// Mock of the hydraulics unit, which is both the brake (I_Brake) and the hydraulics (I_Hydraulics) on MONETS/MONETN.
// The Az/El brake is hydraulic and locks by itself without pressure: Enable := FALSE (hydraulics off) closes the brake, and after
// InjectPressureLoss() the brake is locked and OpenBrake() has no effect until Reset(). Nobody sets Enable TRUE in the rig, so the
// brake opens as before as long as the pressure is there (OpenBrake does not need Enable).
// A close wins over the opening in the same scan, as in HalfBROT FB_HydraulicsControl (a pending bCloseBrake clears bOpenBrake): after
// CloseBrake() an OpenBrake() has no effect until the body has run (the rig calls it at the end of the scan). MONETcommon#272: the
// enabled elevation requests the opening in every scan, after the telescope.
FUNCTION_BLOCK FB_BrakeHydraulicsMock IMPLEMENTS BROTLib.I_Brake, BROTLib.I_Hydraulics
VAR
	bBrakeIsOpen	: BOOL;
	bCloseRequest	: BOOL;	// CloseBrake() in this scan: OpenBrake() is ignored until the body
	bEnabled		: BOOL;
	bFailed			: BOOL;
	bPressureLost	: BOOL;	// InjectPressureLoss: no oil pressure, the brake is locked
	bStartSuction	: BOOL;
	bStopPump		: BOOL;
	nOpenCalls		: UINT;
	nCloseCalls		: UINT;
	nDisableCalls	: UINT;	// Enable := FALSE writes (the hydraulics were switched off)
END_VAR

bCloseRequest := FALSE;	// the scan's close has been applied

METHOD OpenBrake : BOOL
IF NOT bPressureLost AND NOT bCloseRequest THEN
	bBrakeIsOpen := TRUE;
END_IF
nOpenCalls := nOpenCalls + 1;
OpenBrake := NOT bPressureLost;
END_METHOD

METHOD CloseBrake : BOOL
bBrakeIsOpen := FALSE;
bCloseRequest := TRUE;
nCloseCalls := nCloseCalls + 1;
CloseBrake := TRUE;
END_METHOD

// the hydraulics report an error until Reset() (fbHydraulics.Error, #155)
METHOD InjectError
bFailed := TRUE;
END_METHOD

// the hydraulics report an error and the oil pressure is gone: the brake locks at once and cannot be opened until Reset()
// (MonetSafeState_Tests). InjectError alone keeps the pressure (the brake stays as it is).
METHOD InjectPressureLoss
bFailed := TRUE;
bPressureLost := TRUE;
bBrakeIsOpen := FALSE;
END_METHOD

METHOD Reset : BOOL
bFailed := FALSE;
bPressureLost := FALSE;
Reset := TRUE;
END_METHOD

PROPERTY BrakeOpen : BOOL
GET
BrakeOpen := bBrakeIsOpen;
END_GET
END_PROPERTY

PROPERTY Enable : BOOL
GET
Enable := bEnabled;
END_GET
SET
bEnabled := Enable;
IF NOT Enable THEN
	nDisableCalls := nDisableCalls + 1;
	bBrakeIsOpen := FALSE;	// no pressure: the hydraulic brake locks
END_IF
END_SET
END_PROPERTY

PROPERTY Error : BOOL
GET
Error := bFailed;
END_GET
END_PROPERTY

PROPERTY ManualStartSuction : BOOL
GET
ManualStartSuction := bStartSuction;
END_GET
SET
bStartSuction := ManualStartSuction;
END_SET
END_PROPERTY

PROPERTY ManualStopPump : BOOL
GET
ManualStopPump := bStopPump;
END_GET
SET
bStopPump := ManualStopPump;
END_SET
END_PROPERTY

PROPERTY OilPressureOK : BOOL
GET
OilPressureOK := NOT bPressureLost;
END_GET
END_PROPERTY

PROPERTY PumpRunning : BOOL
GET
PumpRunning := bEnabled;
END_GET
END_PROPERTY

PROPERTY SuctionRunning : BOOL
GET
SuctionRunning := FALSE;
END_GET
END_PROPERTY

END_FUNCTION_BLOCK

(* stored: Version 1.1.0.1, ProductVersion 3.1.4024.15
   POU FB_BrakeHydraulicsMock: Id {b710b6cd-5a7f-4296-96e0-69b08cd2bf4f}, SpecialFunc None
   Method OpenBrake: Id {1860ca1d-fc0d-4dcf-9300-461841a019a3}
   Method CloseBrake: Id {c2fadfac-89f8-4739-a96e-c54aa1375935}
   Method InjectError: Id {026406ac-d201-44d8-81fe-06f99e026f89}
   Method InjectPressureLoss: Id {28e89f9d-f339-4cb8-bb99-e89aef723e3b}
   Method Reset: Id {16f43ef0-757d-4384-8dfd-12f9d925c432}
   Property BrakeOpen: Id {204a74e7-dd69-4286-ba4a-f6d8af491b0e}
   Get Get: Id {7906c1ca-cfc4-4697-85f7-4747f39743d8}
   Property Enable: Id {a7fabbdc-1914-4ba3-b880-a9a9efdf711e}
   Get Get: Id {364b7fff-89a5-4852-b599-5d22c51cb154}
   Set Set: Id {8c793db1-1c28-4866-a715-01adc659a592}
   Property Error: Id {279f0a44-7656-4396-a7be-cb44b7e5318c}
   Get Get: Id {4f35eefc-e137-4abb-8542-d2d4aaa06e16}
   Property ManualStartSuction: Id {7f588d9c-ed74-4399-990d-89932edb9a62}
   Get Get: Id {394ff4dd-77fc-4809-923d-7b4194d3838b}
   Set Set: Id {5dd4b46b-9ff7-498a-b2a3-08aecb1c0a0a}
   Property ManualStopPump: Id {2ddff069-acbf-4690-822f-72a1fdad65df}
   Get Get: Id {d181e345-9c59-4ffe-af5d-7f46134ada30}
   Set Set: Id {12230013-e2ae-40c1-8c20-7bb664e59b9b}
   Property OilPressureOK: Id {4e5d1a2f-5061-45bd-afc0-42d65abbac19}
   Get Get: Id {2331e5ef-f7fe-4e8f-bf87-51be9fd5dd72}
   Property PumpRunning: Id {c3c69bdb-57ab-4882-b8ac-0521a24f8c82}
   Get Get: Id {50a048d3-49d3-4e44-a835-795bb82bfb2b}
   Property SuctionRunning: Id {ea33d952-0443-4f26-a4a5-ce0a15f57dca}
   Get Get: Id {82adce1e-1b93-4e60-aecc-0dcb17bd32cf} *)
